(* IEC 61131-3 sources: codesys-to-s7/tests/corpus/C2S7-RING-TODO/neg/input/src/POUs/FB_R, 1 file *)

(* ---- FB_R.decl.st ---- *)
// Автор:      WTP2 (исходный блок S7); перевод в ST — s7conv 0.1.0
// Версия:     1.0 (исходный блок S7)
FUNCTION_BLOCK FB_R
VAR
    a : INT;
    b : INT;
END_VAR
